SUBAPPLICATION OptionalGroup_002 (* Optionsgruppe 2: Digitaler Eingang/Ausgang per Options-Adapter freigeschaltet (QI aus AOption_X_TO_EVENT aktiviert/deaktiviert die ganze Gruppe) *)
  (* Standard: 61499-2; Description: Copyright (c) 2026 Meisterschulen am Ostbahnhof This program and the accompanying materials are made available under the terms of the Eclipse Public License 2.0 which is available at https://www.eclipse.org/legal/epl-2.0/ SPDX-License-Identifier: EPL-2.0 *)
  (* Version 1.0, 2026-10-13, Franz Höpfinger, Meisterschulen am Ostbahnhof *)
  PACKAGE MyLib_AX_Option::sys;
  IMPORT logiBUS::io::DI::logiBUS_DI::Input_I2;
  IMPORT logiBUS::io::DQ::logiBUS_DO::Output_Q2;
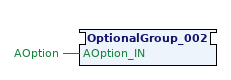
  SOCKETS
    AOption_IN : Option::AOption;
  END_SOCKETS
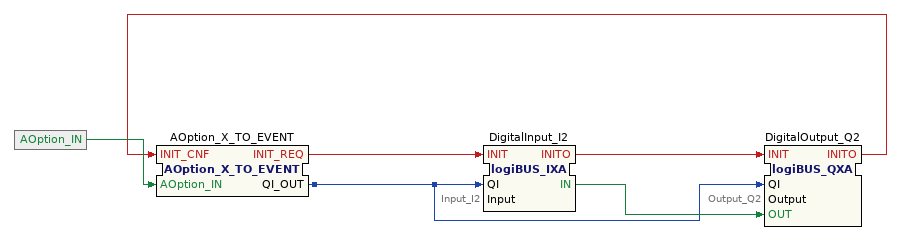
  FBS
    DigitalInput_I2 : logiBUS::io::DI::logiBUS_IXA(Input := Input_I2);
    DigitalOutput_Q2 : logiBUS::io::DQ::logiBUS_QXA(Output := Output_Q2);
    AOption_X_TO_EVENT : Option::conversion::AOption_X_TO_EVENT;
  END_FBS
  EVENT_CONNECTIONS
    AOption_X_TO_EVENT.INIT_REQ TO DigitalInput_I2.INIT;
    DigitalInput_I2.INITO TO DigitalOutput_Q2.INIT;
    DigitalOutput_Q2.INITO TO AOption_X_TO_EVENT.INIT_CNF;
  END_CONNECTIONS
  DATA_CONNECTIONS
    AOption_X_TO_EVENT.QI_OUT TO DigitalInput_I2.QI;
    AOption_X_TO_EVENT.QI_OUT TO DigitalOutput_Q2.QI;
  END_CONNECTIONS
  ADAPTER_CONNECTIONS
    DigitalInput_I2.IN TO DigitalOutput_Q2.OUT;
    AOption_IN TO AOption_X_TO_EVENT.AOption_IN;
  END_CONNECTIONS
END_SUBAPPLICATION
